FUNCTION_BLOCK FB_Gr00Periphery
(*

The function block used to control periphery.

Constructor: 		Patryk Panylo
Company:		E. Riexinger GmbH
Date:			24.10.2015
Version:			1.00

Date:			Revision:		Who:				Comment
dd.mm.yyyy		x.xx			Initials			comment

*)
VAR_INPUT
	(* Input variables / Eingang Variablen *)
	bEnable						:BOOL;						(* Axis present *)
END_VAR
VAR_OUTPUT
	(* Output variables / Ausgang Variablen *)

END_VAR
VAR_IN_OUT
	(* Input Output variables / Ausgang Variablen *)
	Periphery					:FB_PERIPHERY_REF;			(* Interface of periphery *)
END_VAR
VAR
	(* Enummerations *)

	(* Variables *)

	(* References *)

	(* Interfaces *)

	(* Instances *)

END_VAR

IF NOT bEnable								(* Signal FB enable *)
THEN

	RETURN;
END_IF

A_PeripheryLink();

ACTION A_PeripheryLink:

;
END_ACTION

END_FUNCTION_BLOCK

(* stored: Version 1.1.0.1, ProductVersion 3.1.4024.15
   POU FB_Gr00Periphery: Id {31e5a010-d888-4e2b-a250-40e4081ecdd5}, SpecialFunc None
   Action A_PeripheryLink: Id {b7d0f8a2-3b55-4a25-aa80-cfc121469c62} *)
